(* IEC 61131-3 sources: plc-process-lib/tests/POUs/Suites/FB_MotorVfd_Test, 36 files *)

(* ---- CfgChecksRampCommSpeedDevBits.method.decl.st ---- *)
// Переопределение CheckConfig: бит 9 (рампа < 0), бит 10 (tCommLoss = T#0S), бит 11 (rSpeedDev_pct > 0 при
// tSpeedDev = T#0S) и биты FB_Motor вместе (tResetWindow = T#0S — бит 2).
METHOD PRIVATE CfgChecksRampCommSpeedDevBits
VAR
    fbTime    : FB_FakeTime;       // подменное время, старт 1 ч
    fbVfd     : FB_MotorVfd;       // двигатель с ПЧ под тестом
    stCmd     : ST_MotorCmd;       // команды
    stRetain  : ST_DeviceRetain;   // энергонезависимые данные
    stCfg     : ST_MotorCfg;       // конфигурация (умолчания)
    wExpected : WORD;              // ожидаемые биты
END_VAR

(* ---- CommLossCountersFrozen.method.decl.st ---- *)
// ПЧ с ОС из слова состояния работает в Auto 10 с; связь пропала на 1 ч (кабель), питание есть. Через tCommLoss —
// отказ CommLoss, и двигатель больше не считается работающим по устаревшей ОС (VFD-11): xRunning, Running и бит
// RUNNING сняты, наработка выросла только на время до отказа, CurrentRunSeconds = 0. Связь вернулась, ПЧ работает,
// запрос есть — Running без нового пуска.
METHOD PRIVATE CommLossCountersFrozen
VAR
    fbTime   : FB_FakeTime;       // подменное время, старт 1 ч
    fbVfd    : FB_MotorVfd;       // двигатель с ПЧ под тестом
    stCmd    : ST_MotorCmd;       // команды
    stRetain : ST_DeviceRetain;   // энергонезависимые данные
    stCfg    : ST_MotorCfg;       // конфигурация (умолчания)

    udiRun0  : UDINT;             // наработка до потери связи, с
    udiCnt0  : UDINT;             // пусков до потери связи
END_VAR

(* ---- CommLossFaultAfterDelayNotLatched.method.decl.st ---- *)
// Потеря связи (xCommLossIsFault = TRUE): сразу — контроль ОС приостановлен (FB_SUSPENDED), через tCommLoss =
// 3 с — нефиксируемый отказ (бит COMM_LOSS, Fault, выходы сняты, Available = FALSE, тревога слота 6), задание
// удерживается; связь вернулась, ПЧ работает, запрос Auto есть — Running без Reset.
METHOD PRIVATE CommLossFaultAfterDelayNotLatched
VAR
    fbTime   : FB_FakeTime;       // подменное время, старт 1 ч
    fbVfd    : FB_MotorVfd;       // двигатель с ПЧ под тестом
    stCmd    : ST_MotorCmd;       // команды
    stRetain : ST_DeviceRetain;   // энергонезависимые данные
    stCfg    : ST_MotorCfg;       // конфигурация (умолчания)
    itfAlm   : I_Alarm;           // тревога слота
END_VAR

(* ---- CommLossInOosNoFaultNoWarning.method.decl.st ---- *)
// Отказ связи с ПЧ действует во всех режимах, кроме OutOfService (13.6, 14.4): в OOS связи нет 4 с — ни
// MOT_FLT_COMM_LOSS (xCommLossIsFault = TRUE), ни MOT_WRN_COMM_LOSS (FALSE), тревога слота 6 — в OutOfService.
// Выход в Manual при той же потере связи — предупреждение появляется.
METHOD PRIVATE CommLossInOosNoFaultNoWarning
VAR
    fbTime   : FB_FakeTime;       // подменное время, старт 1 ч
    fbVfd    : FB_MotorVfd;       // двигатель с ПЧ под тестом
    stCmd    : ST_MotorCmd;       // команды
    stRetain : ST_DeviceRetain;   // энергонезависимые данные
    stCfg    : ST_MotorCfg;       // конфигурация (умолчания)
    itfAlm   : I_Alarm;           // тревога слота CommLoss
END_VAR

(* ---- CommLossNotFaultWarning.method.decl.st ---- *)
// xCommLossIsFault = FALSE (пуск/стоп и ОС проводами, xFbFromComm = FALSE): потеря связи — только
// предупреждение COMM_LOSS, NE 107 OutOfSpecification и тревога слота 6; двигатель работает, ОС по DI
// контролируется.
METHOD PRIVATE CommLossNotFaultWarning
VAR
    fbTime   : FB_FakeTime;       // подменное время, старт 1 ч
    fbVfd    : FB_MotorVfd;       // двигатель с ПЧ под тестом
    stCmd    : ST_MotorCmd;       // команды
    stRetain : ST_DeviceRetain;   // энергонезависимые данные
    stCfg    : ST_MotorCfg;       // конфигурация (умолчания)
    itfAlm   : I_Alarm;           // тревога слота
END_VAR

(* ---- CommLossSuppressesFeedbackSupervisionImmediately.method.decl.st ---- *)
// Связь пропала во время пуска (tFbStart = 2 с) на 2,4 с — меньше tCommLoss: FailToStart не формируется,
// состояние Starting удерживается; связь вернулась с ОС — Running без отказа.
METHOD PRIVATE CommLossSuppressesFeedbackSupervisionImmediately
VAR
    fbTime   : FB_FakeTime;       // подменное время, старт 1 ч
    fbVfd    : FB_MotorVfd;       // двигатель с ПЧ под тестом
    stCmd    : ST_MotorCmd;       // команды
    stRetain : ST_DeviceRetain;   // энергонезависимые данные
    stCfg    : ST_MotorCfg;       // конфигурация (умолчания)
END_VAR

(* ---- CommLossWhileStoppingHoldsStopping.method.decl.st ---- *)
// Связь с ПЧ пропала во время торможения (Stopping, ОС из слова состояния): ОС недостоверна — состояние
// удерживается в Stopping (не «остановлен»), контроль приостановлен; связь вернулась через 1 с (меньше
// tCommLoss), ПЧ ещё тормозит — Stopping под контролем tFbStop; ПЧ остановился — Stopped без отказа.
METHOD PRIVATE CommLossWhileStoppingHoldsStopping
VAR
    fbTime   : FB_FakeTime;       // подменное время, старт 1 ч
    fbVfd    : FB_MotorVfd;       // двигатель с ПЧ под тестом
    stCmd    : ST_MotorCmd;       // команды
    stRetain : ST_DeviceRetain;   // энергонезависимые данные
    stCfg    : ST_MotorCfg;       // конфигурация (умолчания)
END_VAR

(* ---- CommLostStatusWordIgnored.method.decl.st ---- *)
// Слово состояния ПЧ достоверно только при связи (14.2): связи нет 1 с (меньше tCommLoss), в последнем
// прочитанном слове «авария» и «не готов» — ни ExtFault (дольше tExtFaultFilter), ни PERMIT_MISSING. Связь
// появилась, авария держится — ExtFault через tExtFaultFilter, «не готов» — PERMIT_MISSING.
METHOD PRIVATE CommLostStatusWordIgnored
VAR
    fbTime   : FB_FakeTime;       // подменное время, старт 1 ч
    fbVfd    : FB_MotorVfd;       // двигатель с ПЧ под тестом
    stCmd    : ST_MotorCmd;       // команды
    stRetain : ST_DeviceRetain;   // энергонезависимые данные
    stCfg    : ST_MotorCfg;       // конфигурация (умолчания)
END_VAR

(* ---- CommRestoredRunningWithoutDemandStops.method.decl.st ---- *)
// Manual: отказ связи снимает ручную защёлку; связь вернулась, ПЧ ещё работает, запроса нет — штатный
// останов с контролем (Stopping, команда не подаётся), затем Stopped.
METHOD PRIVATE CommRestoredRunningWithoutDemandStops
VAR
    fbTime   : FB_FakeTime;       // подменное время, старт 1 ч
    fbVfd    : FB_MotorVfd;       // двигатель с ПЧ под тестом
    stCmd    : ST_MotorCmd;       // команды
    stRetain : ST_DeviceRetain;   // энергонезависимые данные
    stCfg    : ST_MotorCfg;       // конфигурация (умолчания)
END_VAR

(* ---- FirstCallFakeTimeCommLossDeterministic.method.decl.st ---- *)
// Связи с ПЧ нет с первого вызова: ResolveTime() до вложенного фильтра даёт подменное время и в первом
// вызове, отказ связи — ровно через tCommLoss = 2 с (на 1,9 с ещё нет).
METHOD PRIVATE FirstCallFakeTimeCommLossDeterministic
VAR
    fbTime   : FB_FakeTime;       // подменное время, старт 1 ч
    fbVfd    : FB_MotorVfd;       // двигатель с ПЧ под тестом
    stCmd    : ST_MotorCmd;       // команды
    stRetain : ST_DeviceRetain;   // энергонезависимые данные
    stCfg    : ST_MotorCfg;       // конфигурация (умолчания)
END_VAR

(* ---- FirstCallSetsTypeMotorVfdAndPassesDefaultCfg.method.decl.st ---- *)
// Чек-лист, пункты 1 и 8: тип MotorVfd (FB_Motor его не затирает), 8 слотов, умолчания Cfg с полем stVfd
// проходят CheckConfig, задание 0 %.
METHOD PRIVATE FirstCallSetsTypeMotorVfdAndPassesDefaultCfg
VAR
    fbTime   : FB_FakeTime;       // подменное время, старт 1 ч
    fbVfd    : FB_MotorVfd;       // двигатель с ПЧ под тестом
    stCmd    : ST_MotorCmd;       // команды
    stRetain : ST_DeviceRetain;   // энергонезависимые данные
    stCfg    : ST_MotorCfg;       // конфигурация (умолчания)
END_VAR

(* ---- ImplementsIMotorPolymorphicArray.method.decl.st ---- *)
// FB_Motor и FB_MotorVfd в одном массиве I_Motor: станция читает Running, Starts, RunSeconds без знания
// типа; тип в stCommon.eDevType — Motor и MotorVfd; Reset() через I_Device.
METHOD PRIVATE ImplementsIMotorPolymorphicArray
VAR
    fbTime         : FB_FakeTime;              // подменное время, старт 1 ч
    fbVfd          : FB_MotorVfd;              // двигатель с ПЧ под тестом
    stCmd          : ST_MotorCmd;              // команды
    stRetain       : ST_DeviceRetain;          // энергонезависимые данные
    stCfg          : ST_MotorCfg;              // конфигурация (умолчания)
    fbTime2        : FB_FakeTime;              // время двигателя прямого пуска
    fbMot          : FB_Motor;                 // двигатель прямого пуска
    stCmd2         : ST_MotorCmd;              // его команды
    stRetain2      : ST_DeviceRetain;          // его энергонезависимые данные
    aitfMot        : ARRAY[1..2] OF I_Motor;   // насосы станции
    itfMot         : I_Motor;                  // насос через интерфейс
    itfDev         : I_Device;                 // устройство через интерфейс
    uiIdx          : UINT;                     // номер насоса
    uiRunningCount : UINT;                     // работающих
    udiStartsSum   : UDINT;                    // пусков всего
    udiRunSum      : UDINT;                    // наработка всего, с
END_VAR

(* ---- ImplementsIMotorPolymorphicArray.method.impl.st ---- *)
coUnit.TEST('MotorVfd_ImplementsIMotor_PolymorphicArray');

fbMot(itfTime := fbTime2, stCmd := stCmd2, stRetain := stRetain2, stCfg := stCfg);
stCmd2.xStart := TRUE;
fbMot.xFbRun := TRUE;
fbTime2.Advance(tStep := T#1S);
fbMot(itfTime := fbTime2, stCmd := stCmd2, stRetain := stRetain2, stCfg := stCfg);
SpinVfd(fbV := fbVfd, fbT := fbTime, stC := stCmd, stR := stRetain, stF := stCfg, uiN := 1, tDt := T#0S);
stCmd.xStart := TRUE;
fbVfd.xVfdRunning := TRUE;
SpinVfd(fbV := fbVfd, fbT := fbTime, stC := stCmd, stR := stRetain, stF := stCfg, uiN := 1, tDt := T#1S);
FOR uiIdx := 1 TO 5 DO
    fbTime2.Advance(tStep := T#1S);
    fbMot(itfTime := fbTime2, stCmd := stCmd2, stRetain := stRetain2, stCfg := stCfg);
END_FOR
SpinVfd(fbV := fbVfd, fbT := fbTime, stC := stCmd, stR := stRetain, stF := stCfg, uiN := 5, tDt := T#1S);
aitfMot[1] := fbMot;
aitfMot[2] := fbVfd;
FOR uiIdx := 1 TO 2 DO
    itfMot := aitfMot[uiIdx];
    IF itfMot.Running THEN
        uiRunningCount := uiRunningCount + 1;
    END_IF
    udiStartsSum := udiStartsSum + itfMot.Starts;
    udiRunSum := udiRunSum + itfMot.RunSeconds;
END_FOR
AssertEquals_UINT(Expected := 2, Actual := uiRunningCount, Message := 'both running via I_Motor');
AssertEquals_UDINT(Expected := 2, Actual := udiStartsSum, Message := 'one start each');
AssertEquals_UDINT(Expected := 10, Actual := udiRunSum, Message := '5 s each');
AssertTrue(Condition := fbMot.stSts.stCommon.eDevType = E_DeviceType.Motor, Message := 'plain motor type');
AssertTrue(Condition := fbVfd.stSts.stCommon.eDevType = E_DeviceType.MotorVfd, Message := 'VFD type');
itfDev := aitfMot[2];
AssertTrue(Condition := itfDev.Reset(), Message := 'Reset via I_Device');

coUnit.TEST_FINISHED();

(* ---- ImplementsIMotorVfdLeadPumpProperties.method.decl.st ---- *)
// I_MotorVfd для ведущего насоса: SpeedRef, SpeedAct, SpeedAutoActive, Running и Mode через интерфейс.
// SpeedAutoActive (VFD-06) — только Auto, Running и без отказа: FALSE у стоящего в Auto насоса, в Starting (ОС ещё
// нет), в Stopping (ОС ещё есть), при отказе связи и в Manual; TRUE — Auto и Running.
METHOD PRIVATE ImplementsIMotorVfdLeadPumpProperties
VAR
    fbTime   : FB_FakeTime;       // подменное время, старт 1 ч
    fbVfd    : FB_MotorVfd;       // двигатель с ПЧ под тестом
    stCmd    : ST_MotorCmd;       // команды
    stRetain : ST_DeviceRetain;   // энергонезависимые данные
    stCfg    : ST_MotorCfg;       // конфигурация (умолчания)
    itfLead  : I_MotorVfd;        // ведущий насос через интерфейс
END_VAR

(* ---- InvalidSpeedLimitsCfgErrBit8.method.decl.st ---- *)
// Пределы скорости неверны (min >= max, max > 100, min < 0): бит 8 MOT_CFG_VFD_SPEED_LIMITS (переопределение
// CheckConfig вызывается и из тела FB_Motor), CheckFunction.
METHOD PRIVATE InvalidSpeedLimitsCfgErrBit8
VAR
    fbTime   : FB_FakeTime;       // подменное время, старт 1 ч
    fbVfd    : FB_MotorVfd;       // двигатель с ПЧ под тестом
    stCmd    : ST_MotorCmd;       // команды
    stRetain : ST_DeviceRetain;   // энергонезависимые данные
    stCfg    : ST_MotorCfg;       // конфигурация (умолчания)
END_VAR

(* ---- LocalModeRefTracksActualSpeed.method.decl.st ---- *)
// Local: выходы сняты, задание и задание оператора следят за фактической скоростью (42 %); возврат в Manual
// при работающем ПЧ — без рывка задания.
METHOD PRIVATE LocalModeRefTracksActualSpeed
VAR
    fbTime   : FB_FakeTime;       // подменное время, старт 1 ч
    fbVfd    : FB_MotorVfd;       // двигатель с ПЧ под тестом
    stCmd    : ST_MotorCmd;       // команды
    stRetain : ST_DeviceRetain;   // энергонезависимые данные
    stCfg    : ST_MotorCfg;       // конфигурация (умолчания)
END_VAR

(* ---- ManualSpeedTracksAutoForBumpless.method.decl.st ---- *)
// В Auto задание оператора следит за целью (60 %); переход в Manual — задание не прыгает, команда работы
// сохраняется.
METHOD PRIVATE ManualSpeedTracksAutoForBumpless
VAR
    fbTime   : FB_FakeTime;       // подменное время, старт 1 ч
    fbVfd    : FB_MotorVfd;       // двигатель с ПЧ под тестом
    stCmd    : ST_MotorCmd;       // команды
    stRetain : ST_DeviceRetain;   // энергонезависимые данные
    stCfg    : ST_MotorCfg;       // конфигурация (умолчания)
END_VAR

(* ---- PlcRestartCommLaterAdoptedWithoutFault.method.decl.st ---- *)
// Старт ПЛК, ПЧ работает, ОС — из слова состояния, но связи первые 0,5 с нет (мастер Modbus ещё не опросил
// слейв): подхват ждёт первой достоверной ОС — при появлении связи двигатель подхвачен (Running, команда), без
// UncommandedRun и без счёта пуска.
METHOD PRIVATE PlcRestartCommLaterAdoptedWithoutFault
VAR
    fbTime   : FB_FakeTime;       // подменное время, старт 1 ч
    fbVfd    : FB_MotorVfd;       // двигатель с ПЧ под тестом
    stCmd    : ST_MotorCmd;       // команды
    stRetain : ST_DeviceRetain;   // энергонезависимые данные
    stCfg    : ST_MotorCfg;       // конфигурация (умолчания)
END_VAR

(* ---- PlcRestartFbFromDiAdoptedWithoutFault.method.decl.st ---- *)
// Старт ПЛК, ОС по DI (xFbFromComm = FALSE), слово состояния ПЧ ещё не прочитано: в первом вызове точки
// расширения берут корректную stCfg, а не умолчания — двигатель подхвачен, UncommandedRun нет.
METHOD PRIVATE PlcRestartFbFromDiAdoptedWithoutFault
VAR
    fbTime   : FB_FakeTime;       // подменное время, старт 1 ч
    fbVfd    : FB_MotorVfd;       // двигатель с ПЧ под тестом
    stCmd    : ST_MotorCmd;       // команды
    stRetain : ST_DeviceRetain;   // энергонезависимые данные
    stCfg    : ST_MotorCfg;       // конфигурация (умолчания)
END_VAR

(* ---- PlcRestartRefBumpless.method.decl.st ---- *)
// Перезапуск ПЛК при работающем ПЧ: подхват (VFD-09). Auto, запрос есть, ПЧ на 70 %: задание на ПЧ сразу 70 % —
// фактическая скорость в пределах rSpeedMin…rSpeedMax, — без провала к 0 и рампы с нуля (rRampUp 10 %/с). Manual,
// ПЧ на 55 %: подхват пишет фактическую скорость и в задание оператора stCmd.rSpeedSp_pct (оно не энергонезависимо
// и после старта 0) — двигатель не тормозится до rSpeedMin.
METHOD PRIVATE PlcRestartRefBumpless
VAR
    fbTime   : FB_FakeTime;       // подменное время, старт 1 ч
    fbVfd    : FB_MotorVfd;       // двигатель с ПЧ под тестом
    stCmd    : ST_MotorCmd;       // команды
    stRetain : ST_DeviceRetain;   // энергонезависимые данные
    stCfg    : ST_MotorCfg;       // конфигурация (умолчания)

    fbTime2  : FB_FakeTime;       // время второго двигателя
    fbVfd2   : FB_MotorVfd;       // двигатель в Manual
    stCmd2   : ST_MotorCmd;       // его команды
    stRet2   : ST_DeviceRetain;   // его данные (Manual)
END_VAR

(* ---- PowerLossCommLossNoFaultNotRunning.method.decl.st ---- *)
// Пропало питание станции: xPowerOk = FALSE, ПЧ обесточен, связи нет (VFD-11, VFD-12). Отказа CommLoss и тревоги
// слота 6 нет — пропадание питания — останов без отказа (13.7); двигатель не работает: xRunning снят сразу,
// Stopped, наработка за час не растёт. Питание вернулось — ПЧ загружается VFD_POWER_UP_DELAY = 10 с, затем фильтр
// tCommLoss = 3 с: отказ связи — только через 13 с, если связь так и не появилась; связь есть — отказ снят.
METHOD PRIVATE PowerLossCommLossNoFaultNotRunning
VAR
    fbTime   : FB_FakeTime;       // подменное время, старт 1 ч
    fbVfd    : FB_MotorVfd;       // двигатель с ПЧ под тестом
    stCmd    : ST_MotorCmd;       // команды
    stRetain : ST_DeviceRetain;   // энергонезависимые данные
    stCfg    : ST_MotorCfg;       // конфигурация (умолчания)

    udiRun0  : UDINT;             // наработка до пропадания питания, с
    itfAlm   : I_Alarm;           // тревога слота CommLoss
END_VAR

(* ---- SlowRamp1msCycleNotStalled.method.decl.st ---- *)
// Рампа задания 0,003 %/с при цикле 1 мс (VFD-13): состояние рампы в LREAL — за 1 с задание растёт на 0,003 %
// (в REAL приращение 3·10⁻⁶ % рядом с 70 % терялось бы и рампа стояла). Ожидаемое: 70 + 0,003 · 1 с.
METHOD PRIVATE SlowRamp1msCycleNotStalled
VAR
    fbTime   : FB_FakeTime;       // подменное время, старт 1 ч
    fbVfd    : FB_MotorVfd;       // двигатель с ПЧ под тестом
    stCmd    : ST_MotorCmd;       // команды
    stRetain : ST_DeviceRetain;   // энергонезависимые данные
    stCfg    : ST_MotorCfg;       // конфигурация (умолчания)
END_VAR

(* ---- SpeedActNaNStsFinite.method.decl.st ---- *)
// Фактическая скорость NaN при xCommOk (мусор Modbus): связь недостоверна, задание удерживается; в Sts и свойстве
// SpeedAct — конечное 0.0 (R6: карта регистров NaN не получает).
METHOD PRIVATE SpeedActNaNStsFinite
VAR
    fbTime   : FB_FakeTime;       // подменное время, старт 1 ч
    fbVfd    : FB_MotorVfd;       // двигатель с ПЧ под тестом
    stCmd    : ST_MotorCmd;       // команды
    stRetain : ST_DeviceRetain;   // энергонезависимые данные
    stCfg    : ST_MotorCfg;       // конфигурация (умолчания)

    uBits    : U_RealBits;        // NaN по битам
    itfLead  : I_MotorVfd;        // двигатель через интерфейс
END_VAR

(* ---- SpeedClampedToMinMax.method.decl.st ---- *)
// Пределы задания 20…90 %: цель Auto 95 % → 90 % (слежение stCmd.rSpeedSp_pct тоже 90), 5 % → 20 %;
// в Manual 150 % → 90 % и записывается обратно в stCmd.
METHOD PRIVATE SpeedClampedToMinMax
VAR
    fbTime   : FB_FakeTime;       // подменное время, старт 1 ч
    fbVfd    : FB_MotorVfd;       // двигатель с ПЧ под тестом
    stCmd    : ST_MotorCmd;       // команды
    stRetain : ST_DeviceRetain;   // энергонезависимые данные
    stCfg    : ST_MotorCfg;       // конфигурация (умолчания)
END_VAR

(* ---- SpeedDeviationDuringRampIgnored.method.decl.st ---- *)
// Рассогласование во время рампы не контролируется: рост 1 %/с к цели 50 %, факт отстаёт (0 %) — за 20 с
// (больше tSpeedDev = 2 с при допуске 10 %) предупреждения нет (задание 20 %); рампа завершена — предупреждение
// ровно через tSpeedDev. Источник: tools/reference/motor.py, сценарий ramp_slow_20s.
METHOD PRIVATE SpeedDeviationDuringRampIgnored
VAR
    fbTime   : FB_FakeTime;       // подменное время, старт 1 ч
    fbVfd    : FB_MotorVfd;       // двигатель с ПЧ под тестом
    stCmd    : ST_MotorCmd;       // команды
    stRetain : ST_DeviceRetain;   // энергонезависимые данные
    stCfg    : ST_MotorCfg;       // конфигурация (умолчания)
END_VAR

(* ---- SpeedDeviationWarningAfterDelay.method.decl.st ---- *)
// Рассогласование задания 50 % и факта 35 % (больше rSpeedDev_pct = 10 %) дольше tSpeedDev = 10 с:
// предупреждение SPEED_DEV, NE 107 OutOfSpecification, тревога слота 7; не отказ — двигатель работает.
METHOD PRIVATE SpeedDeviationWarningAfterDelay
VAR
    fbTime   : FB_FakeTime;       // подменное время, старт 1 ч
    fbVfd    : FB_MotorVfd;       // двигатель с ПЧ под тестом
    stCmd    : ST_MotorCmd;       // команды
    stRetain : ST_DeviceRetain;   // энергонезависимые данные
    stCfg    : ST_MotorCfg;       // конфигурация (умолчания)
    itfAlm   : I_Alarm;           // тревога слота
END_VAR

(* ---- SpeedRampLimitsRate.method.decl.st ---- *)
// Рампа задания: min 20 %, рост 10 %/с, спад 5 %/с, шаг 100 мс; пуск — с 20 %, через 1,5 с — 35 %, через 3 с —
// цель 50 %; цель 30 %: через 2 с — 40 %, через 4 с — 30 %. Источник: tools/reference/motor.py, сценарии ramp_*.
METHOD PRIVATE SpeedRampLimitsRate
VAR
    fbTime   : FB_FakeTime;       // подменное время, старт 1 ч
    fbVfd    : FB_MotorVfd;       // двигатель с ПЧ под тестом
    stCmd    : ST_MotorCmd;       // команды
    stRetain : ST_DeviceRetain;   // энергонезависимые данные
    stCfg    : ST_MotorCfg;       // конфигурация (умолчания)
END_VAR

(* ---- SpeedSpNaNHoldsRef.method.decl.st ---- *)
// Цель не конечна (NaN от ПИД/Modbus): задание удерживается, предупреждение SPEED_SP_INVALID, NaN в задание
// оператора не пишется; конечная цель снова принимается.
METHOD PRIVATE SpeedSpNaNHoldsRef
VAR
    fbTime   : FB_FakeTime;       // подменное время, старт 1 ч
    fbVfd    : FB_MotorVfd;       // двигатель с ПЧ под тестом
    stCmd    : ST_MotorCmd;       // команды
    stRetain : ST_DeviceRetain;   // энергонезависимые данные
    stCfg    : ST_MotorCfg;       // конфигурация (умолчания)
    uBits    : U_RealBits;        // NaN по битам
END_VAR

(* ---- SpinVfd.method.decl.st ---- *)
// Помощник: uiN вызовов двигателя с ПЧ, перед каждым — шаг подменного времени tDt (T#0S — тот же момент).
// Входы тест пишет по имени экземпляра до вызова помощника; ассертов внутри нет
METHOD PRIVATE SpinVfd
VAR_IN_OUT
    fbV : FB_MotorVfd;       // двигатель с ПЧ
    fbT : FB_FakeTime;       // подменное время
    stC : ST_MotorCmd;       // команды
    stR : ST_DeviceRetain;   // энергонезависимые данные
END_VAR
VAR_IN_OUT CONSTANT
    stF : ST_MotorCfg;       // конфигурация
END_VAR
VAR_INPUT
    uiN : UINT;              // число вызовов
    tDt : TIME;              // шаг времени перед каждым вызовом
END_VAR
VAR
    uiLoop : UINT;           // номер вызова
END_VAR

(* ---- SpinVfd.method.impl.st ---- *)
FOR uiLoop := 1 TO uiN DO
    fbT.Advance(tStep := tDt);
    fbV(itfTime := fbT, stCmd := stC, stRetain := stR, stCfg := stF);
END_FOR

(* ---- StartInCommGapRefPresetToMin.method.decl.st ---- *)
// Пуск в Manual во время короткого пропуска связи (короче tCommLoss): пуск не блокируется, а задание передать
// нельзя — предустановка rSpeedMin ждёт связи (VFD-10). Связь вернулась — задание 30 % (rSpeedMin), а не рампа от
// 0; дальше рампа 1 %/с: 30,1 % через 0,1 с.
METHOD PRIVATE StartInCommGapRefPresetToMin
VAR
    fbTime   : FB_FakeTime;       // подменное время, старт 1 ч
    fbVfd    : FB_MotorVfd;       // двигатель с ПЧ под тестом
    stCmd    : ST_MotorCmd;       // команды
    stRetain : ST_DeviceRetain;   // энергонезависимые данные
    stCfg    : ST_MotorCfg;       // конфигурация (умолчания)
END_VAR

(* ---- StartPresetsRampToMin.method.decl.st ---- *)
// Вход в Starting начинает рампу с rSpeedMin_pct = 30 % (а не с 0): в вызове пуска 30 %, через шаг 100 мс —
// 31 %, через 1 с — 40 % (рост 10 %/с, цель 80 %). Источник: tools/reference/motor.py, сценарии start_preset_*.
METHOD PRIVATE StartPresetsRampToMin
VAR
    fbTime   : FB_FakeTime;       // подменное время, старт 1 ч
    fbVfd    : FB_MotorVfd;       // двигатель с ПЧ под тестом
    stCmd    : ST_MotorCmd;       // команды
    stRetain : ST_DeviceRetain;   // энергонезависимые данные
    stCfg    : ST_MotorCfg;       // конфигурация (умолчания)
END_VAR

(* ---- StartWithNaNTargetRefStartsAtMin.method.decl.st ---- *)
// Пуск при не конечной цели (ПИД выдал NaN, пока насос стоял), без ограничения роста (rRampUp_pctps = 0):
// задание начинается с rSpeedMin_pct = 25 %, а не с последней конечной цели 60 %; предупреждение
// SPEED_SP_INVALID. Конечная цель — задание сразу к ней (VFD-03).
METHOD PRIVATE StartWithNaNTargetRefStartsAtMin
VAR
    fbTime   : FB_FakeTime;       // подменное время, старт 1 ч
    fbVfd    : FB_MotorVfd;       // двигатель с ПЧ под тестом
    stCmd    : ST_MotorCmd;       // команды
    stRetain : ST_DeviceRetain;   // энергонезависимые данные
    stCfg    : ST_MotorCfg;       // конфигурация
    uBits    : U_RealBits;        // NaN по битам
END_VAR

(* ---- StopSetsRefZero.method.decl.st ---- *)
// «Стоп» снимает команду работы и задание — 0 % в том же вызове (торможение — рампой ПЧ).
METHOD PRIVATE StopSetsRefZero
VAR
    fbTime   : FB_FakeTime;       // подменное время, старт 1 ч
    fbVfd    : FB_MotorVfd;       // двигатель с ПЧ под тестом
    stCmd    : ST_MotorCmd;       // команды
    stRetain : ST_DeviceRetain;   // энергонезависимые данные
    stCfg    : ST_MotorCfg;       // конфигурация (умолчания)
END_VAR

(* ---- VfdFaultTripsAndResetPulses.method.decl.st ---- *)
// Авария ПЧ из слова состояния — внешняя авария (фильтр 200 мс, фиксируется); Reset даёт импульс xQReset,
// ПЧ сбрасывает аварию через 0,5 с — отказ снят в окне без второго нажатия.
METHOD PRIVATE VfdFaultTripsAndResetPulses
VAR
    fbTime   : FB_FakeTime;       // подменное время, старт 1 ч
    fbVfd    : FB_MotorVfd;       // двигатель с ПЧ под тестом
    stCmd    : ST_MotorCmd;       // команды
    stRetain : ST_DeviceRetain;   // энергонезависимые данные
    stCfg    : ST_MotorCfg;       // конфигурация (умолчания)
END_VAR

(* ---- VfdNotReadyBlocksStart.method.decl.st ---- *)
// ПЧ не готов (xVfdReady = FALSE при связи): пуск оператора — RejectedPermit, бит PERMIT_MISSING; в Auto запрос
// ждёт (ReadyToStart = FALSE) и пуск происходит, когда ПЧ готов.
METHOD PRIVATE VfdNotReadyBlocksStart
VAR
    fbTime   : FB_FakeTime;       // подменное время, старт 1 ч
    fbVfd    : FB_MotorVfd;       // двигатель с ПЧ под тестом
    stCmd    : ST_MotorCmd;       // команды
    stRetain : ST_DeviceRetain;   // энергонезависимые данные
    stCfg    : ST_MotorCfg;       // конфигурация (умолчания)
END_VAR
